(* IEC 61131-3 sources: rusty/tests/lit/single/oop, 33 files *)

(* ---- aggregate_return_complex.st ---- *)
// RUN: %COMPILE %s && %RUN | %CHECK %s
FUNCTION_BLOCK fb_with_method
VAR_TEMP
    ret : ARRAY[0..1] OF STRING;
    ret_struct : returnStruct;
END_VAR
    METHOD method_with_aggregagte_return: ARRAY[0..1] OF STRING
    VAR_INPUT
        in: STRING;
        in2: STRING;
    END_VAR
        method_with_aggregagte_return[0] := in;
        method_with_aggregagte_return[1] := in2;
    END_METHOD

    METHOD method_with_struct_return: returnStruct
    VAR_INPUT
        in: STRING;
        in2: STRING;
    END_VAR
       method_with_struct_return.a := in;
       method_with_struct_return.b := in2;

       method_with_struct_return.c[0][0] := 'a';
       method_with_struct_return.c[0][1] := 'b';
       method_with_struct_return.c[1][0] := 'c';
       method_with_struct_return.c[1][1] := 'd';
    END_METHOD

    ret := method_with_aggregagte_return('Hello', 'World!');
    printf('%s$N', ADR(ret[0])); // CHECK: Hello
    printf('%s$N', ADR(ret[1])); // CHECK: World!

    ret_struct := method_with_struct_return('Hello', 'Again!');
    printf('%s$N', ADR(ret_struct.a)); // CHECK: Hello
    printf('%s$N', ADR(ret_struct.b)); // CHECK: Again!

    printf('%s$N', ADR(ret_struct.c[0][0])); // CHECK: a
    printf('%s$N', ADR(ret_struct.c[0][1])); // CHECK: b
    printf('%s$N', ADR(ret_struct.c[1][0])); // CHECK: c
    printf('%s$N', ADR(ret_struct.c[1][1])); // CHECK: d
END_FUNCTION_BLOCK

FUNCTION main
VAR
    fb: fb_with_method;
    ret : ARRAY[0..1] OF STRING;
    ret_struct : returnStruct;
END_VAR
    fb();
    ret := fb.method_with_aggregagte_return('Goodbye', 'World!');
    printf('%s$N', ADR(ret[0])); // CHECK: Goodbye
    printf('%s$N', ADR(ret[1])); // CHECK: World!
    ret_struct := fb.method_with_struct_return('Goodbye', 'Again!');
    printf('%s$N', ADR(ret_struct.a)); // CHECK: Goodbye
    printf('%s$N', ADR(ret_struct.b)); // CHECK: Again!
    printf('%s$N', ADR(ret_struct.c[0][0])); // CHECK: a
    printf('%s$N', ADR(ret_struct.c[0][1])); // CHECK: b
    printf('%s$N', ADR(ret_struct.c[1][0])); // CHECK: c
    printf('%s$N', ADR(ret_struct.c[1][1])); // CHECK: d
END_FUNCTION

TYPE returnStruct : STRUCT
    a : STRING;
    b : STRING;
    c : ARRAY[0..1] OF ARRAY[0..1] OF STRING;
END_STRUCT
END_TYPE

(* ---- aggregate_return_types.st ---- *)
// RUN: %COMPILE %s && %RUN | %CHECK %s
FUNCTION_BLOCK fb_with_method
VAR_TEMP
    ret : STRING;
END_VAR
    METHOD method_with_aggregagte_return: STRING
    VAR_INPUT
        in: STRING;
    END_VAR
        method_with_aggregagte_return := in;
    END_METHOD

    ret := method_with_aggregagte_return('Hello');
    printf('%s$N', ADR(ret)); // CHECK: Hello
END_FUNCTION_BLOCK

FUNCTION main
VAR
    fb: fb_with_method;
    ret : STRING;
END_VAR

    fb();
    ret := fb.method_with_aggregagte_return('World!');
    printf('%s$N', ADR(ret)); // CHECK: World!
END_FUNCTION

(* ---- fb_access_members_from_base.st ---- *)
// RUN: %COMPILE %s && %RUN | %CHECK %s
FUNCTION_BLOCK fb
VAR
    x : INT;
    y : INT;
END_VAR
END_FUNCTION_BLOCK

FUNCTION_BLOCK fb2 EXTENDS fb
END_FUNCTION_BLOCK

FUNCTION_BLOCK foo
VAR
    myFb : fb2;
END_VAR
    myFb.x := 1;
    printf('%d$N', myFb.x); //CHECK: 1
END_FUNCTION_BLOCK

FUNCTION main : DINT
    VAR
        fb :foo;
    END_VAR
    fb();
END_FUNCTION

(* ---- fb_complex_access_of_super_members.st ---- *)
// RUN: %COMPILE %s && %RUN | %CHECK %s
FUNCTION_BLOCK grandparent
VAR
    y : ARRAY[0..5] OF INT;
    a : INT;
END_VAR
END_FUNCTION_BLOCK

FUNCTION_BLOCK parent extends grandparent
    VAR
        x : ARRAY[0..10] OF INT;
        b : INT;
    END_VAR
END_FUNCTION_BLOCK

FUNCTION_BLOCK child EXTENDS parent
    VAR
        z : ARRAY[0..10] OF INT;
    END_VAR
    y[b + z[b*2] - a] := 20;
    b := 1;
    z[b] := 3;
    z[b*2] := 4;
    a := 2;
    y[b + z[b*2] - a] := 60;
    printf('%d$N', y[0]); //CHECK: 20
    printf('%d$N', y[3]); //CHECK: 60
END_FUNCTION_BLOCK

FUNCTION main : DINT
    VAR
        fb : child;
    END_VAR
    fb();
END_FUNCTION

(* ---- fb_direct_calls.st ---- *)
// RUN: %COMPILE %s && %RUN | %CHECK %s

TYPE Position2D:
    STRUCT
        x: DINT;
        y: DINT;
    END_STRUCT
END_TYPE

TYPE Position3D:
    STRUCT
        x: DINT;
        y: DINT;
        z: DINT;
    END_STRUCT
END_TYPE

FUNCTION_BLOCK FbA
    VAR
        placeholderA: STRING;
    END_VAR

    VAR_INPUT
        x: DINT;
        y: DINT;
    END_VAR

    VAR_OUTPUT
        result2D: Position2D;
    END_VAR

    result2D.x := x;
    result2D.y := y;
END_FUNCTION_BLOCK

FUNCTION_BLOCK FbB EXTENDS FbA
    VAR_INPUT
        z: DINT;
    END_VAR

    VAR_OUTPUT
        result3D: Position3D;
    END_VAR

    // using the values from FbA
    result3D.x := x;
    result3D.y := y;
    result3D.z := z;
END_FUNCTION_BLOCK

FUNCTION_BLOCK FbC EXTENDS FbB
    VAR_INPUT
        multiplier2D: DINT;
        multiplier3D: DINT;
    END_VAR

    VAR
        placeholderC1: STRING;
        placeholderC2: INT;
    END_VAR

    VAR_IN_OUT
        resultMultiplied2D: Position2D;
        resultMultiplied3D: Position3D;
    END_VAR

    resultMultiplied2D.x := x * multiplier2D;
    resultMultiplied2D.y := y * multiplier2D;

    resultMultiplied3D.x := x * multiplier3D;
    resultMultiplied3D.y := y * multiplier3D;
    resultMultiplied3D.z := z * multiplier3D;
END_FUNCTION_BLOCK

FUNCTION main
    VAR
        instanceA: FbA;
        instanceB: FbB;
        instanceC: FbC;

        pos2D: Position2D;
        pos3D: Position3D;
    END_VAR

    // CHECK: Position2D(10, 20)
    instanceA(
        x := 10,
        result2D => pos2D,
        y := 20,
    );
    printf('Position2D(%d, %d)$N', pos2D.x, pos2D.y);

    // CHECK-NEXT: Position3D(40, 50, 60)
    instanceB(
        z := 60,
        y := 50,
        result3D => pos3D,
        x := 40,
    );
    printf('Position3D(%d, %d, %d)$N', pos3D.x, pos3D.y, pos3D.z);

    // CHECK-NEXT: Position2D(140, 160)
    // CHECK-NEXT: Position3D(280, 320, 360)
    instanceC(
        multiplier2D := 2,
        z := 90,
        x := 70,
        resultMultiplied3D := pos3D,
        y := 80,
        multiplier3D := 4,
        resultMultiplied2D := pos2D,
    );
    printf('Position2D(%d, %d)$N', pos2D.x, pos2D.y);
    printf('Position3D(%d, %d, %d)$N', pos3D.x, pos3D.y, pos3D.z);
END_FUNCTION

(* ---- fb_init_at_both_levels_runs_once.st ---- *)
// RUN: %COMPILE %s && %RUN | %CHECK %s
// Regression: when both Base and Child declare `FB_INIT`, each must run
// exactly once during construction. Pre-fix the doubled base-ctor (issue 1)
// and the inherited FB_INIT re-emit (issue 2) inflated these counts.
FUNCTION_BLOCK Base
VAR
    base_calls : DINT := 0;
END_VAR
    METHOD FB_INIT
        base_calls := base_calls + 1;
    END_METHOD
END_FUNCTION_BLOCK

FUNCTION_BLOCK Child EXTENDS Base
VAR
    child_calls : DINT := 0;
END_VAR
    METHOD FB_INIT
        child_calls := child_calls + 1;
    END_METHOD
END_FUNCTION_BLOCK

FUNCTION main : DINT
VAR
    c : Child;
END_VAR
    printf('%d$N', c.base_calls);  // CHECK: 1
    printf('%d$N', c.child_calls); // CHECK: 1
END_FUNCTION

(* ---- fb_init_base_runs_before_child.st ---- *)
// RUN: %COMPILE %s && %RUN | %CHECK %s
// Sequencing: `Base.FB_INIT` must run before `Child.FB_INIT`, so that the
// child's body can rely on initialized base state. Pre-fix, the doubled base
// ctor would still produce the right value here, but the inherited-FB_INIT
// re-emit ran the base FB_INIT after derived members were touched, which
// could clobber values written by the child. We pin the post-fix order.
FUNCTION_BLOCK Base
VAR
    x : DINT := 0;
END_VAR
    METHOD FB_INIT
        x := 10;
    END_METHOD
END_FUNCTION_BLOCK

FUNCTION_BLOCK Child EXTENDS Base
VAR
    y : DINT := 0;
END_VAR
    METHOD FB_INIT
        // Base.FB_INIT must have already run, so x == 10 here.
        y := x * 2;
    END_METHOD
END_FUNCTION_BLOCK

FUNCTION main : DINT
VAR
    c : Child;
END_VAR
    printf('%d$N', c.x); // CHECK: 10
    printf('%d$N', c.y); // CHECK: 20
END_FUNCTION

(* ---- fb_init_inherited_runs_once.st ---- *)
// RUN: %COMPILE %s && %RUN | %CHECK %s
// Regression: an inherited `FB_INIT` must only run once per construction.
// Pre-fix the derived ctor invoked it both via the base ctor chain and via a
// spurious second emit (find_method walked up the super class).
FUNCTION_BLOCK Base
VAR
    init_calls : DINT := 0;
END_VAR
    METHOD FB_INIT
        init_calls := init_calls + 1;
    END_METHOD
END_FUNCTION_BLOCK

FUNCTION_BLOCK Child EXTENDS Base
END_FUNCTION_BLOCK

FUNCTION main : DINT
VAR
    c : Child;
END_VAR
    printf('%d$N', c.init_calls); // CHECK: 1
END_FUNCTION

(* ---- fb_init_runs_per_instance.st ---- *)
// RUN: %COMPILE %s && %RUN | %CHECK %s
// Sanity: the fix for double base-ctor / inherited FB_INIT must not
// over-correct. Each constructed instance must still run the inherited
// `FB_INIT` once. Two instances => count of 2.
VAR_GLOBAL
    base_init_count : DINT := 0;
END_VAR

FUNCTION_BLOCK Base
    METHOD FB_INIT
        base_init_count := base_init_count + 1;
    END_METHOD
END_FUNCTION_BLOCK

FUNCTION_BLOCK Child EXTENDS Base
END_FUNCTION_BLOCK

FUNCTION main : DINT
VAR
    a : Child;
    b : Child;
END_VAR
    printf('%d$N', base_init_count); // CHECK: 2
END_FUNCTION

(* ---- fb_method_callled.st ---- *)
// RUN: %COMPILE %s && %RUN | %CHECK %s
FUNCTION_BLOCK foo
VAR
    bar: DINT := 42;
END_VAR
    METHOD addToBar: DINT
    VAR_INPUT
        in: INT;
    END_VAR
        bar := in + bar;
        addToBar := bar;
    END_METHOD

    addToBar(3);
    printf('%d$N', bar); // CHECK: 45
END_FUNCTION_BLOCK

FUNCTION main
VAR
    fb: foo;
    x: DINT;
END_VAR
    fb();
    x := fb.addToBar(3);
    printf('%d$N', x); // CHECK: 48
END_FUNCTION

(* ---- fb_method_shadowing.st ---- *)
// RUN: %COMPILE %s && %RUN | %CHECK %s
FUNCTION_BLOCK foo
VAR
    bar: DINT := 42;
END_VAR
    METHOD addToBar: DINT
    VAR_INPUT
        in: INT;
    END_VAR
    VAR
        bar: DINT := 17;
    END_VAR
        bar := in + bar;
        addToBar := bar;
    END_METHOD
    METHOD addToLocalBar: DINT
    VAR_INPUT
        in: INT;
    END_VAR
    VAR
        bar: DINT := 17;
    END_VAR
        this^.bar := in + bar;
        addToLocalBar := this^.bar;
    END_METHOD

    addToBar(3);
    printf('%d$N', bar); // CHECK: 42
END_FUNCTION_BLOCK

FUNCTION main
VAR
    fb: foo;
    x: DINT;
END_VAR
    fb();
    x := fb.addToBar(3);
    printf('%d$N', x); // CHECK: 20
    x := fb.addToLocalBar(46);
    printf('%d$N', x); // CHECK: 63
END_FUNCTION

(* ---- fb_method_with_explicit_return.st ---- *)
// RUN: %COMPILE %s && %RUN | %CHECK %s
FUNCTION_BLOCK fb
    METHOD foo : STRING
        VAR_INPUT
            x : DINT;
        END_VAR
        foo := 'hello';
    END_METHOD
END_FUNCTION_BLOCK
FUNCTION main : DINT
VAR
    my_fb : fb;
    res : STRING;
END_VAR
    res := my_fb.foo(x := 1);
    printf('%s$N', ADR(res)); // CHECK: hello
END_FUNCTION

(* ---- fb_with_in_and_out_extension.st ---- *)
// RUN: %COMPILE %s && %RUN | %CHECK %s
FUNCTION_BLOCK foo
METHOD met1 : INT
    VAR_INPUT
    mandatoryInput : INT;
    optionalInput : INT := 5;
    END_VAR
    VAR_OUTPUT
    outputValue : INT;
    END_VAR
    outputValue := mandatoryInput + optionalInput;
    printf('method 1 - mandatoryInput: %d, optionalInput: %d$N', mandatoryInput, optionalInput);
END_METHOD
END_FUNCTION_BLOCK

FUNCTION_BLOCK foo2 EXTENDS foo
VAR
    x : INT;
END_VAR
met1(
	mandatoryInput := 0,
	optionalInput := 0,
	outputValue => x
);
// CHECK: method 1 - mandatoryInput: 0, optionalInput: 0
// CHECK: method output : 0
printf('method output : %d$N', x);
met1(
	mandatoryInput := 5,
	outputValue => x
);
// CHECK: method 1 - mandatoryInput: 5, optionalInput: 5
// CHECK: method output : 10
printf('method output : %d$N', x);
END_FUNCTION_BLOCK

FUNCTION main : DINT
VAR
    foo_inst: foo;
    foo2_inst : foo2;
    out : INT;
END_VAR
foo2_inst();

foo_inst.met1(mandatoryInput:= 2, outputValue => out);
// CHECK: method 1 - mandatoryInput: 2, optionalInput: 5
// CHECK: method output : 7
printf('method output : %d$N', out);

foo2_inst.met1(mandatoryInput:= 1, outputValue => out);
// CHECK: method 1 - mandatoryInput: 1, optionalInput: 5
// CHECK: method output : 6
printf('method output : %d$N', out);

END_FUNCTION

(* ---- fb_with_super_class_method_calls.st ---- *)
// RUN: %COMPILE %s && %RUN | %CHECK %s
FUNCTION_BLOCK foo
VAR
    s : STRING;
END_VAR
METHOD baz
    s := 'hello';
END_METHOD
END_FUNCTION_BLOCK

FUNCTION_BLOCK bar EXTENDS foo
    s := 'world';
END_FUNCTION_BLOCK

FUNCTION main: DINT
VAR
    fb: bar;
END_VAR
    fb.baz();
    printf('%s$N', REF(fb.s)); // CHECK: hello
    fb();
    printf('%s$N', REF(fb.s)); // CHECK: world
END_FUNCTION

(* ---- grandparent_access_through_super.st ---- *)
// RUN: %COMPILE %s && %RUN | %CHECK %s
FUNCTION_BLOCK grandparent
VAR
    x : INT := 10;
END_VAR
END_FUNCTION_BLOCK

FUNCTION_BLOCK parent EXTENDS grandparent
VAR
    y : INT := 20;
END_VAR
END_FUNCTION_BLOCK

FUNCTION_BLOCK child EXTENDS parent
    // Access parent member directly with SUPER^
    SUPER^.y := 100;
    // Access grandparent member through SUPER^
    SUPER^.x := 200;
END_FUNCTION_BLOCK

FUNCTION main
VAR
    c : child;
END_VAR
    c();
    // Check if the values are set correctly
    printf('%d$N', c.x); // CHECK: 200
    printf('%d$N', c.y); // CHECK: 100
END_FUNCTION

(* ---- method_call_through_struct_field.st ---- *)
// RUN: %COMPILE %s && %RUN | %CHECK %s

// Anchors that a chained qualified call (`h.inst.bar()`) resolves end-to-end
// when the call's operator is a multi-level ReferenceExpr whose base is itself
// a ReferenceExpr. Counterpart to the resolver-only unit test
// `chained_qualified_call_resolves_through_recursive_bases`.
FUNCTION_BLOCK SomeFb
    METHOD bar : INT
        bar := 7;
    END_METHOD
END_FUNCTION_BLOCK

TYPE Holder : STRUCT inst : SomeFb; END_STRUCT END_TYPE

FUNCTION main : DINT
    VAR
        h : Holder;
        x : INT;
    END_VAR

    x := h.inst.bar();
    printf('chained=%d$N', x);
    // CHECK: chained=7
END_FUNCTION

(* ---- method_initial_values.st ---- *)
// RUN: %COMPILE %s && %RUN | %CHECK %s
FUNCTION_BLOCK MyClass
    VAR
        x, y : INT;
    END_VAR

    METHOD testMethod
    VAR_INPUT
        myMethodArg : INT := 3;
    END_VAR
        x := myMethodArg;
    END_METHOD
END_FUNCTION_BLOCK

FUNCTION main
VAR
cl : MyClass;
END_VAR
    cl.testMethod();
    printf('%d$N', cl.x); // CHECK: 3
END_FUNCTION

(* ---- method_var_output.st ---- *)
// RUN: %COMPILE %s && %RUN | %CHECK %s
FUNCTION_BLOCK foo
METHOD baz
VAR_OUTPUT
    out : STRING;
END_VAR
    out := 'hello';
END_METHOD
END_FUNCTION_BLOCK

FUNCTION main
VAR
    s: STRING;
    fb: foo;
END_VAR
    fb.baz(out => s);
    printf('%s$n', REF(s)); // CHECK: hello
    s := 'reset';
    printf('%s$n', REF(s)); // CHECK: reset
    fb.baz(s);
    printf('%s$n', REF(s)); // CHECK: hello
END_FUNCTION

(* ---- parent_variable_access_in_method.st ---- *)
// RUN: %COMPILE %s && %RUN | %CHECK %s
FUNCTION_BLOCK foo
    VAR
        x: DINT := 50;
    END_VAR
END_FUNCTION_BLOCK

FUNCTION_BLOCK bar EXTENDS foo
    METHOD set0 // TODO(volsa): https://github.com/PLC-lang/rusty/issues/1408
        x := 25;
    END_METHOD

    METHOD shadowed
    VAR
        x: DINT := 100;
    END_VAR
    END_METHOD
END_FUNCTION_BLOCK

FUNCTION main
    VAR
        instance: bar;
    END_VAR

    instance.set0();
    printf('%d$N', instance.x); // CHECK: 25
    // assigning to a locally shadowed variable should not change the parent variable
    instance.shadowed();
    printf('%d$N', instance.x); // CHECK: 25
END_FUNCTION

(* ---- super_basic_access.st ---- *)
// RUN: %COMPILE %s && %RUN | %CHECK %s
FUNCTION_BLOCK parent
VAR
    x : INT := 10;
    y : INT := 20;
END_VAR

METHOD get_sum : INT
    get_sum := x + y;
END_METHOD
END_FUNCTION_BLOCK

FUNCTION_BLOCK child EXTENDS parent
METHOD get_values : INT
    VAR
        x : INT := 100; // Shadows parent's x
    END_VAR
    VAR_INPUT
        use_parent : BOOL;
    END_VAR

    IF use_parent THEN
        get_values := SUPER^.x + y; // Use parent's x but child inherits y
    ELSE
        get_values := x + y; // Use shadowed x and inherited y
    END_IF;
END_METHOD

    printf('x = %d$N', x);                          // CHECK: x = 10
    printf('SUPER^.x = %d$N', SUPER^.x);            // CHECK: SUPER^.x = 10
    printf('y = %d$N', y);                          // CHECK: y = 20
    printf('get_values(TRUE) = %d$N', get_values(TRUE));    // CHECK: get_values(TRUE) = 30
    printf('get_values(FALSE) = %d$N', get_values(FALSE));  // CHECK: get_values(FALSE) = 120
    printf('SUPER^.get_sum() = %d$N', SUPER^.get_sum());    // CHECK: SUPER^.get_sum() = 30
END_FUNCTION_BLOCK

FUNCTION main : INT
VAR
    inst : child;
END_VAR
    inst();
END_FUNCTION

(* ---- super_constant_in_initializer.st ---- *)
// RUN: %COMPILE %s && %RUN | %CHECK %s
FUNCTION_BLOCK grandparent
VAR CONSTANT
    base_value : INT := 42;
END_VAR
END_FUNCTION_BLOCK

FUNCTION_BLOCK parent EXTENDS grandparent
END_FUNCTION_BLOCK

FUNCTION_BLOCK child EXTENDS parent
VAR CONSTANT
    const_from_super : INT := SUPER^.base_value + 1;
END_VAR
VAR
    var_from_super : INT := SUPER^.base_value;
    var_from_inherited : INT := base_value * 2;
END_VAR
VAR_TEMP
    temp_from_super : INT := SUPER^.base_value;
END_VAR
    printf('const_from_super = %d$N', const_from_super);        // CHECK: const_from_super = 43
    printf('var_from_super = %d$N', var_from_super);            // CHECK: var_from_super = 42
    printf('var_from_inherited = %d$N', var_from_inherited);    // CHECK: var_from_inherited = 84
    printf('temp_from_super = %d$N', temp_from_super);          // CHECK: temp_from_super = 42
END_FUNCTION_BLOCK

FUNCTION main : INT
VAR
    inst : child;
END_VAR
    inst();
END_FUNCTION

(* ---- super_in_control_structures.st ---- *)
// RUN: %COMPILE %s && %RUN | %CHECK %s
FUNCTION_BLOCK parent
VAR
    counter : INT := 0;
    threshold : INT := 5;
END_VAR

METHOD increment : INT
    counter := counter + 1;
    increment := counter;
END_METHOD

METHOD reset
    counter := 0;
END_METHOD
END_FUNCTION_BLOCK

FUNCTION_BLOCK child EXTENDS parent
METHOD increment : INT
    increment := SUPER^.increment() + 1; // Increment parent's counter and add 1
END_METHOD
METHOD test
    VAR
        i : INT;
        result : INT;
    END_VAR

    // Reset parent's counter
    SUPER^.reset();

    // Use SUPER^ in IF statement
    // CHECK: Initial counter: 0
    IF SUPER^.counter < SUPER^.threshold THEN
        printf('Initial counter: %d$N', SUPER^.counter);
    END_IF;

    // Use SUPER^ in FOR loop
    // CHECK: Loop increment: 1
    // CHECK: Loop increment: 2
    // CHECK: Loop increment: 3
    FOR i := 1 TO 3 BY 1 DO
        result := SUPER^.increment();
        printf('Loop increment: %d$N', result);
    END_FOR;

    // Use SUPER^ in CASE statement
    CASE SUPER^.counter OF
        // CHECK: Counter is three
        3: printf('Counter is three$N');
        4: printf('Counter is four$N');
    END_CASE;

    // Use SUPER^ in WHILE loop
    // CHECK: While increment: 4
    // CHECK: While increment: 5
    WHILE SUPER^.counter < 5 DO
        result := SUPER^.increment();
        printf('While increment: %d$N', result);
    END_WHILE;
END_METHOD

    test();

    // CHECK: Parent counter: 5
    printf('Parent counter: %d$N', SUPER^.counter);
END_FUNCTION_BLOCK

FUNCTION main : INT
VAR
    inst : child;
END_VAR
    inst();
END_FUNCTION

(* ---- super_keyword_overridden_method.st ---- *)
// RUN: %COMPILE %s && %RUN | %CHECK %s
FUNCTION_BLOCK fb
VAR
    x: INT := 10;
END_VAR

METHOD foo : INT
    VAR_INPUT
        a: INT := 100;
    END_VAR

    foo := a + x;
END_METHOD
END_FUNCTION_BLOCK

FUNCTION_BLOCK fb2 EXTENDS fb
// TODO: should shadowing parent variables with temp vars be allowed?
// uncommenting the following var-block will cause a compile error
// VAR_TEMP
//     x: INT := 20;
// END_VAR
METHOD foo : INT
    VAR_INPUT
        a: INT := 1000;
    END_VAR

    foo := a - x;
END_METHOD

    printf('%d$N', super^.foo(super^.x));   // CHECK: 20
    printf('%d$N', super^.foo(x));          // CHECK: 20
    printf('%d$N', super^.foo());           // CHECK: 110
    printf('%d$N', foo(super^.x));          // CHECK: 0
    printf('%d$N', foo(x));                 // CHECK: 0
    printf('%d$N', foo());                  // CHECK: 990
END_FUNCTION_BLOCK

FUNCTION main
VAR
    inst: fb2;
END_VAR
    inst();
END_FUNCTION

(* ---- super_multi_level_inheritance.st ---- *)
// RUN: %COMPILE %s && %RUN | %CHECK %s
FUNCTION_BLOCK grandparent
VAR
    gp_value : INT := 100;
END_VAR

METHOD calculate : INT
    calculate := gp_value;
END_METHOD
END_FUNCTION_BLOCK

FUNCTION_BLOCK parent EXTENDS grandparent
VAR
    p_value : INT := 200;
END_VAR

METHOD calculate : INT
    calculate := p_value + SUPER^.calculate();
END_METHOD
END_FUNCTION_BLOCK

FUNCTION_BLOCK child EXTENDS parent
VAR
    c_value : INT := 300;
END_VAR

METHOD calculate : INT
    calculate := c_value + SUPER^.calculate();
END_METHOD

    // Access values from different levels
    printf('c_value = %d$N', c_value);                // CHECK: c_value = 300
    printf('p_value = %d$N', p_value);                // CHECK: p_value = 200
    printf('gp_value = %d$N', gp_value);              // CHECK: gp_value = 100

    // Call methods from different inheritance levels
    printf('calculate() = %d$N', calculate());        // CHECK: calculate() = 600
    printf('SUPER^.calculate() = %d$N', SUPER^.calculate());  // CHECK: SUPER^.calculate() = 300
END_FUNCTION_BLOCK

FUNCTION main : INT
VAR
    inst : child;
END_VAR
    inst();
END_FUNCTION

(* ---- super_with_parenthesized_expressions.st ---- *)
// RUN: %COMPILE %s && %RUN | %CHECK %s
FUNCTION_BLOCK parent
VAR
    x: INT := 10;
    y: INT := 20;
    z: INT := 30;
END_VAR

METHOD calculate: INT
    VAR_INPUT
        a: INT;
        b: INT;
    END_VAR
    calculate := a * b;
END_METHOD

METHOD get_value: INT
    get_value := x + y + z;
END_METHOD
END_FUNCTION_BLOCK

FUNCTION_BLOCK child EXTENDS parent
VAR
    multiplier: INT := 3;
END_VAR

METHOD test
    VAR
        result: INT;
    END_VAR

    // Basic parenthesized expression with SUPER
    result := (SUPER^.x + SUPER^.y);
    // CHECK: Basic parentheses: 30
    printf('Basic parentheses: %d$N', result);

    // Nested parentheses with SUPER
    result := ((SUPER^.x + SUPER^.y) * (SUPER^.z));
    // CHECK: Nested parentheses: 900
    printf('Nested parentheses: %d$N', result);

    // Parenthesized expression with method call
    result := (SUPER^.x + SUPER^.y + (SUPER^.calculate(SUPER^.x, SUPER^.y)));
    // CHECK: Expression with method: 230
    printf('Expression with method: %d$N', result);

    // Complex calculation with mixed precedence and parentheses
    result := ((SUPER^.x * multiplier) + (SUPER^.y * 2) + SUPER^.z);
    // CHECK: Complex calculation: 100
    printf('Complex calculation: %d$N', result);

    // Conditional expression with parentheses
    IF ((SUPER^.x + SUPER^.y) > SUPER^.z) THEN
        result := 42;
    ELSE
        result := 24;
    END_IF;
    // CHECK: Conditional with parentheses: 24
    printf('Conditional with parentheses: %d$N', result);

    // Combined SUPER references across parentheses
    result := (SUPER^.get_value()) + (SUPER^.x * SUPER^.y / 2);
    // CHECK: Combined SUPER references: 160
    printf('Combined SUPER references: %d$N', result);
END_METHOD

END_FUNCTION_BLOCK

FUNCTION main: INT
VAR
    inst: child;
END_VAR
    inst.test();
END_FUNCTION

(* ---- super_without_deref.st ---- *)
// RUN: %COMPILE %s && %RUN | %CHECK %s
FUNCTION_BLOCK parent
VAR
    value : INT := 42;
END_VAR

METHOD get_value : INT
    get_value := value;
END_METHOD
END_FUNCTION_BLOCK

FUNCTION_BLOCK child EXTENDS parent
VAR
    p_ref : REF_TO parent;
END_VAR

    // SUPER without deref creates a reference
    p_ref := SUPER;

    // Accessing through reference
    printf('p_ref^.value = %d$N', p_ref^.value);      // CHECK: p_ref^.value = 42
    printf('p_ref^.get_value() = %d$N', p_ref^.get_value()); // CHECK: p_ref^.get_value() = 42

    // Modifying through reference
    p_ref^.value := 100;
    printf('SUPER^.value after modification = %d$N', SUPER^.value); // CHECK: SUPER^.value after modification = 100

    // Compare direct access vs reference access
    printf('Are they equal? %d$N', SUPER^.value = p_ref^.value); // CHECK: Are they equal? 1
END_FUNCTION_BLOCK

FUNCTION main : INT
VAR
    inst : child;
END_VAR
    inst();
END_FUNCTION

(* ---- this_basic_access.st ---- *)
// RUN: %COMPILE %s && %RUN | %CHECK %s
FUNCTION_BLOCK fb
VAR
    x : INT := 10;
    y : INT := 20;
END_VAR

METHOD get_sum : INT
    get_sum := x + y;
END_METHOD
METHOD get_values : INT
    VAR
        x : INT := 100; // Shadows fb's x
        y : INT := 200; // Shadows fb's y
    END_VAR
    VAR_INPUT
        use_function_block : BOOL;
    END_VAR

    IF use_function_block THEN
        get_values := THIS^.x + y; // Use fb's x but local y
    ELSE
        get_values := x + y; // Use shadowed x and y
    END_IF;
END_METHOD

    printf('x = %d$N', x);                          // CHECK: x = 10
    printf('THIS^.x = %d$N', THIS^.x);            // CHECK: THIS^.x = 10
    printf('y = %d$N', y);                          // CHECK: y = 20
    printf('get_values(TRUE) = %d$N', get_values(TRUE));    // CHECK: get_values(TRUE) = 210
    printf('get_values(FALSE) = %d$N', get_values(FALSE));  // CHECK: get_values(FALSE) = 300
    printf('THIS^.get_sum() = %d$N', THIS^.get_sum());    // CHECK: THIS^.get_sum() = 30
END_FUNCTION_BLOCK

FUNCTION main : INT
VAR
    inst : fb;
END_VAR

    inst();
END_FUNCTION

(* ---- this_in_control_structures.st ---- *)
// RUN: %COMPILE %s && %RUN | %CHECK %s
FUNCTION_BLOCK child
VAR
    counter : INT := 0;
    threshold : INT := 5;
END_VAR

METHOD increment : INT
    counter := counter + 1;
    increment := counter;
END_METHOD

METHOD reset
    counter := 0;
END_METHOD
METHOD test
    VAR
        i : INT;
        result : INT;
    END_VAR

    // Reset parent's counter
    THIS^.reset();

    // Use THIS^ in IF statement
    // CHECK: Initial counter: 0
    IF THIS^.counter < THIS^.threshold THEN
        printf('Initial counter: %d$N', THIS^.counter);
    END_IF;

    // Use THIS^ in FOR loop
    // CHECK: Loop increment: 1
    // CHECK: Loop increment: 2
    // CHECK: Loop increment: 3
    FOR i := 1 TO 3 BY 1 DO
        result := THIS^.increment();
        printf('Loop increment: %d$N', result);
    END_FOR;

    // Use THIS^ in CASE statement
    CASE THIS^.counter OF
        // CHECK: Counter is three
        3: printf('Counter is three$N');
        4: printf('Counter is four$N');
    END_CASE;

    // Use THIS^ in WHILE loop
    // CHECK: While increment: 4
    // CHECK: While increment: 5
    WHILE THIS^.counter < 5 DO
        result := THIS^.increment();
        printf('While increment: %d$N', result);
    END_WHILE;
END_METHOD

    test();

    // CHECK: Parent counter: 5
    printf('Parent counter: %d$N', THIS^.counter);
END_FUNCTION_BLOCK

FUNCTION main : INT
VAR
    inst : child;
END_VAR
    inst();
END_FUNCTION

(* ---- this_member_access_without_deref_errors.st ---- *)
// RUN: rm -f %t.out
// RUN: not %COMPILE --error-format clang %s 2>&1 | %CHECK %s
// RUN: test ! -e %t.out

// Regression test for #1728: `THIS.<member>` without an explicit `^` deref
// must be rejected by validation, not silently passed through to codegen
// (where it used to crash with "GEP pointee is not a struct").

// CHECK: {{.*}}this_member_access_without_deref_errors.st:{{[0-9]+}}:{{[0-9]+}}:{{.*}}error[E141]: Cannot access `a` on `POINTER TO fb`; dereference with `^` first
// CHECK: error: Compilation aborted due to critical errors

INTERFACE IAnimal
    METHOD legs : DINT
    END_METHOD
END_INTERFACE

FUNCTION_BLOCK fb
VAR
    a : IAnimal;
END_VAR
METHOD m : DINT
    THIS.a.legs();
END_METHOD
END_FUNCTION_BLOCK

(* ---- this_with_parenthesized_expressions.st ---- *)
// RUN: %COMPILE %s && %RUN | %CHECK %s
FUNCTION_BLOCK fb
VAR
    multiplier: INT := 3;
    x: INT := 10;
    y: INT := 20;
    z: INT := 30;
END_VAR

METHOD calculate: INT
    VAR_INPUT
        a: INT;
        b: INT;
    END_VAR
    calculate := a * b;
END_METHOD

METHOD get_value: INT
    get_value := x + y + z;
END_METHOD

METHOD test
    VAR
        result: INT;
    END_VAR

    // Basic parenthesized expression with THIS
    result := (THIS^.x + THIS^.y);
    // CHECK: Basic parentheses: 30
    printf('Basic parentheses: %d$N', result);

    // Nested parentheses with THIS
    result := ((THIS^.x + THIS^.y) * (THIS^.z));
    // CHECK: Nested parentheses: 900
    printf('Nested parentheses: %d$N', result);

    // Parenthesized expression with method call
    result := (THIS^.x + THIS^.y + (THIS^.calculate(THIS^.x, THIS^.y)));
    // CHECK: Expression with method: 230
    printf('Expression with method: %d$N', result);

    // Complex calculation with mixed precedence and parentheses
    result := ((THIS^.x * multiplier) + (THIS^.y * 2) + THIS^.z);
    // CHECK: Complex calculation: 100
    printf('Complex calculation: %d$N', result);

    // Conditional expression with parentheses
    IF ((THIS^.x + THIS^.y) > THIS^.z) THEN
        result := 42;
    ELSE
        result := 24;
    END_IF;
    // CHECK: Conditional with parentheses: 24
    printf('Conditional with parentheses: %d$N', result);

    // Combined THIS references across parentheses
    result := (THIS^.get_value()) + (THIS^.x * THIS^.y / 2);
    // CHECK: Combined THIS references: 160
    printf('Combined THIS references: %d$N', result);
END_METHOD

END_FUNCTION_BLOCK

FUNCTION main: INT
VAR
    inst: fb;
END_VAR
    inst.test();
END_FUNCTION

(* ---- this_without_deref.st ---- *)
// RUN: %COMPILE %s && %RUN | %CHECK %s
FUNCTION_BLOCK fb
VAR
    p_ref : REF_TO fb;
    value : INT := 42;
END_VAR

METHOD get_value : INT
get_value := value;
END_METHOD

    // THIS without deref creates a reference
    p_ref := THIS;

    // Accessing through reference
    printf('p_ref^.value = %d$N', p_ref^.value);      // CHECK: p_ref^.value = 42
    printf('p_ref^.get_value() = %d$N', p_ref^.get_value()); // CHECK: p_ref^.get_value() = 42

    // Modifying through reference
    p_ref^.value := 100;
    printf('THIS^.value after modification = %d$N', THIS^.value); // CHECK: THIS^.value after modification = 100

    // Compare direct access vs reference access
    printf('Are they equal? %d$N', THIS^.value = p_ref^.value); // CHECK: Are they equal? 1
END_FUNCTION_BLOCK

FUNCTION main : INT
VAR
    inst : fb;
END_VAR
    inst();
END_FUNCTION

(* ---- program_method_called.st ---- *)
// RUN: %COMPILE %s && %RUN | %CHECK %s
PROGRAM foo
VAR
    bar: DINT := 42;
END_VAR
    METHOD addToBar: DINT
    VAR_INPUT
        in: INT;
    END_VAR
        bar := in + bar;
        addToBar := bar;
    END_METHOD

    addToBar(3);
    printf('%d$N', bar); // CHECK: 45
END_PROGRAM

FUNCTION main
VAR
    x: DINT;
END_VAR
    foo();
    x := foo.addToBar(3);
    printf('%d$N', x); // CHECK: 48
END_FUNCTION

(* ---- program_method_shadowing.st ---- *)
// RUN: %COMPILE %s && %RUN | %CHECK %s
PROGRAM foo
VAR
    bar: DINT := 42;
END_VAR
    METHOD addToBar: DINT
    VAR_INPUT
        in: INT;
    END_VAR
    VAR
        bar: DINT := 17;
    END_VAR
        bar := in + bar;
        addToBar := bar;
    END_METHOD

    addToBar(3);
    printf('%d$N', bar); // CHECK: 42
END_PROGRAM

FUNCTION main
VAR
    x: DINT;
END_VAR
    foo();
    x := foo.addToBar(3);
    printf('%d$N', x); // CHECK: 20
END_FUNCTION
